TYPE ST_EL3356ChannelState_1 :
STRUCT
	bOverrange				:BOOL;			(* State Overrange *)
	bDataInvalid				:BOOL;			(* State Data invalid *)
	bError 					:BOOL;			(* State error *)
	bCalibrationInProgress 	:BOOL;			(* State calibration in progress *)
	bSteadyState 			:BOOL;			(* Stady state *)
	bSyncError				:BOOL;			(* Sync error *)
	bToggle					:BOOL;			(* TxPDO Toggle *)
END_STRUCT
END_TYPE

(* stored: Version 1.1.0.1, ProductVersion 3.1.4024.15
   DUT ST_EL3356ChannelState_1: Id {9bbfe096-b05d-4a61-bb45-abd4832c956a} *)
